# EPICS substitutions: iocs/motor/pi-ioc/db/PI_C862.substitutions
# C's iocPI PI_C862.substitutions, P and C from st.cmd.
#
# PI C-862/C-863: one motor record for the controller's single axis, DTYP
# "PIC862" with OUT #C$(C) S0.
file "$(MOTOR)/db/motor.db"
{
pattern
{N,  M,        DTYP,      S,  DESC,          EGU,      DIR,  VELO,  VBAS,  ACCL,  BDST,  BVEL,  BACC,  MRES,  PREC,  DHLM,  DLLM,  INIT}
{3,  "m$(N)",  "PIC862",  0,  "motor $(N)",  degrees,  Pos,  1,     .1,    .2,    0,     1,     .2,    0.01,  5,     100,   -100,  ""}
}
